// TIA Portal V20 export
// export: Created 2026-10-19T18:02:19.6646874Z, ExportSetting WithDefaults, DisplayName Totally Integrated Automation Portal, DisplayVersion V20 Update 6, DisplayName TIA Portal Openness, DisplayVersion V20 Update 6, DisplayName TIA Portal Version Control Interface, DisplayVersion V20 Update 6, DisplayName SINAMICS Startdrive Advanced, DisplayVersion V20 SP1, DisplayName SINAMICS Startdrive G130, G150, S120, S150, SINAMICS MV, G220, S200, S210, DisplayVersion V20 SP1, DisplayName SINAMICS Startdrive G110M, G120, G120C, G120D, G120P, G115D, DisplayVersion V20 SP1, DisplayName STEP 7 Professional, DisplayVersion V20 Update 6, DisplayName STEP 7 Safety, DisplayVersion V20 Update 2, DisplayName WinCC Basic/Comfort/Advanced, DisplayVersion V20 Update 6, DisplayName WinCC Unified, DisplayVersion V20 Update 6
FUNCTION "OUTPUTS" : Void   // FC5, SCL
{ S7_Optimized_Access := 'TRUE' }
VERSION : 0.1
// stored: AutoNumber true, IsIECCheckEnabled false, SetENOAutomatically false, UDAEnableTagReadback false
BEGIN

   // Let's do it for each Shuttle 
   //IF destinationid = position id = id charger (*Setpoint in the HMI reggarding to the charger position*)
   //     2000 = 2000 = 2000 // Example 1 Shuttle on charger positio => Charger on
   //     2000 = 1900 = 2000 // Example 2 Shuttle in other position => Charger off
   //     1000 = 2000 = 2000 // Example 3 Shuttle in charger position but received an order to move to other position => Charger off
   // Enable the charger (Variable) = TRUE;
   //ELSE  
     // Disable the charger
     // Enable the charger (Variable) = FALSE;
   //END_IF;


   IF "FirstScan" THEN
       "Charger Panel" := TRUE;
   END_IF;

   "Charger Panel" := "Charger";

   "Pick Station light" := "Control_DB".Pick_Station.PushButtonLight;
END_FUNCTION
